// TIA Portal V19 export
// export: Created 2026-10-15T10:10:35.0325176Z, ExportSetting WithDefaults, DisplayName Totally Integrated Automation Portal, DisplayVersion V19, DisplayName TIA Portal Openness, DisplayVersion V19, DisplayName TIA Portal Version Control Interface, DisplayVersion V19, DisplayName STEP 7 Professional, DisplayVersion V19, DisplayName STEP 7 Safety, DisplayVersion V19, DisplayName WinCC Basic/Comfort/Advanced, DisplayVersion V19, DisplayName WinCC Unified, DisplayVersion V19
FUNCTION "ROLL_FB69" : Void   // FC10, SCL
{ S7_Optimized_Access := 'TRUE' }
VERSION : 0.1
// stored: AutoNumber true, IsIECCheckEnabled false, SetENOAutomatically false, UDAEnableTagReadback false
BEGIN

   IF "ROLL_State".M[240, 0] AND "ROLL_State".M[240, 1] THEN
       "ROLL_SetMWord"(FirstByte := 240,
                       Value := W#16#2005);
   ELSE
       "ROLL_SetMWord"(FirstByte := 240,
                       Value := W#16#1005);
   END_IF;
END_FUNCTION
